TYPE ST_Prod_Param_Stirrer :
STRUCT
	Mode		: E_Stirrer_mode;
	Speed		: REAL:=1200;
	Flip_mode	: BOOL;
	tON			: INT:=10;	//minutes
	tOFF		: INT:=2;	//minutes


END_STRUCT
END_TYPE

(* stored: Version 1.1.0.1, ProductVersion 3.1.4024.15
   DUT ST_Prod_Param_Stirrer: Id {0798f669-897a-4685-88a7-40bb95aef99f} *)
